Fanuc KAREL source: kt00403.KL

-- PROVISIONAL review KL for V940-1; original PC SHA256 ab83fb77827297d08b7cd990723ab987200e26a5fc27d66088cf6b0e6752b8d5
-- Incomplete behavior may be omitted. Consult companion uncertainty JSON. Do not deploy.
PROGRAM KT00403
%NOLOCKGROUP
VAR
  I1 : INTEGER
  OUT : BOOLEAN
-- UNRESOLVED_DECL Y2 type=002018
BEGIN
  -- V9_ZERO_TABLE_METADATA_HINT layout=0001; no indexed target words; source/name/runtime held
  -- UNRESOLVED_PC offsets 5-16; opcodes 2E,23
  -- UNRESOLVED_PC offsets 21-35; opcodes 2E,22,9D,33,B2
  -- UNRESOLVED_PC offsets 40-62; opcodes 21,22,9D,33,B1,5B,23
  -- UNRESOLVED_PC offsets 67-71; opcodes 7F
END KT00403
